(* IEC 61131-3 sources: Digital-Twin/picode/digital-twin-device/openPLC_v3/webserver/st_files (part 2) *)

(* ---- 924959.st ---- *)
TYPE
  datatype0 : BOOL;
END_TYPE

PROGRAM my_first_program
  VAR
    temp AT %IW1.0 : INT;
    out AT %QW0.0 : INT;
  END_VAR
  VAR
    sp : REAL := 1376.0;
    x0 : REAL := 0.0;
    tr : REAL := 0.001;
    td : REAL := 50.0;
    kp : REAL := 0.00005;
    PID0 : PID;
    GT39_OUT : BOOL;
    INT_TO_REAL28_OUT : REAL;
    REAL_TO_INT34_OUT : INT;
  END_VAR

  GT39_OUT := GT(temp, 1200);
  INT_TO_REAL28_OUT := INT_TO_REAL(temp);
  PID0(AUTO := GT39_OUT, PV := INT_TO_REAL28_OUT, SP := sp, X0 := x0, KP := kp, TR := tr, TD := td, CYCLE := T#1s);
  REAL_TO_INT34_OUT := REAL_TO_INT(PID0.XOUT);
  out := REAL_TO_INT34_OUT;
END_PROGRAM

CONFIGURATION Config0

  RESOURCE Res0 ON PLC
    TASK mytask(INTERVAL := T#50ms,PRIORITY := 0);
    PROGRAM my WITH mytask : my_first_program;
  END_RESOURCE
END_CONFIGURATION

(* ---- 925603.st ---- *)
TYPE
  datatype0 : BOOL;
END_TYPE

PROGRAM my_first_program
  VAR
    temp AT %IW1.0 : INT;
    out AT %QW0.0 : INT;
  END_VAR
  VAR
    sp : REAL := 1030.0;
    x0 : REAL := 0.0;
    tr : REAL := 0.001;
    td : REAL := 50.0;
    kp : REAL := 0.00005;
    PID0 : PID;
    GT39_OUT : BOOL;
    INT_TO_REAL28_OUT : REAL;
    REAL_TO_INT34_OUT : INT;
  END_VAR

  GT39_OUT := GT(temp, 1040);
  INT_TO_REAL28_OUT := INT_TO_REAL(temp);
  PID0(AUTO := GT39_OUT, PV := INT_TO_REAL28_OUT, SP := sp, X0 := x0, KP := kp, TR := tr, TD := td, CYCLE := T#1s);
  REAL_TO_INT34_OUT := REAL_TO_INT(PID0.XOUT);
  out := REAL_TO_INT34_OUT;
END_PROGRAM

CONFIGURATION Config0

  RESOURCE Res0 ON PLC
    TASK mytask(INTERVAL := T#50ms,PRIORITY := 0);
    PROGRAM my WITH mytask : my_first_program;
  END_RESOURCE
END_CONFIGURATION

(* ---- 926092.st ---- *)
PROGRAM my_first_program
  VAR
    temp AT %IW0.0 : INT;
    lamp AT %QX0.0 : BOOL;
    lamp1 AT %QX0.2 : BOOL;
  END_VAR
  VAR
    GT7_OUT : BOOL;
    GT1_OUT : BOOL;
  END_VAR

  GT7_OUT := GT(temp, 17170);
  lamp := GT7_OUT;
  GT1_OUT := GT(temp, 18350);
  lamp1 := GT1_OUT;
END_PROGRAM

CONFIGURATION Config0

  RESOURCE Res0 ON PLC
    TASK mytask(INTERVAL := T#50ms,PRIORITY := 0);
    PROGRAM my WITH mytask : my_first_program;
  END_RESOURCE
END_CONFIGURATION

(* ---- 939656.st ---- *)
PROGRAM my_first_program
  VAR
    temp AT %IW0.0 : INT;
    lamp AT %QX0.0 : BOOL;
    lamp1 AT %QX0.2 : BOOL;
  END_VAR
  VAR
    GT7_OUT : BOOL;
    GT1_OUT : BOOL;
  END_VAR

  GT7_OUT := GT(temp, 17170);
  lamp := GT7_OUT;
  GT1_OUT := GT(temp, 18350);
  lamp1 := GT1_OUT;
END_PROGRAM

CONFIGURATION Config0

  RESOURCE Res0 ON PLC
    TASK mytask(INTERVAL := T#50ms,PRIORITY := 0);
    PROGRAM my WITH mytask : my_first_program;
  END_RESOURCE
END_CONFIGURATION

(* ---- 953895.st ---- *)
PROGRAM program0
  VAR
    PID0 : PID;
    Kp : REAL := 0.01;
    Ki : REAL := 0.1;
    Kd : REAL := 50.0;
  END_VAR
  VAR
    Temperature AT %IW1 : UINT;
    Flow AT %QW0 : UINT;
  END_VAR
  VAR
    Setpoint : UINT := 2500;
    Zero : REAL := 0.0;
    GT13_OUT : BOOL;
    UINT_TO_REAL1_OUT : REAL;
    UINT_TO_REAL9_OUT : REAL;
    REAL_TO_UINT11_OUT : UINT;
  END_VAR

  GT13_OUT := GT(Temperature, Setpoint);
  UINT_TO_REAL1_OUT := UINT_TO_REAL(Temperature);
  UINT_TO_REAL9_OUT := UINT_TO_REAL(Setpoint);
  PID0(AUTO := GT13_OUT, PV := UINT_TO_REAL1_OUT, SP := UINT_TO_REAL9_OUT, X0 := Zero, KP := Kp, TR := Ki, TD := Kd, CYCLE := T#50ms);
  REAL_TO_UINT11_OUT := REAL_TO_UINT(PID0.XOUT);
  Flow := REAL_TO_UINT11_OUT;
END_PROGRAM

CONFIGURATION Config0

  RESOURCE Res0 ON PLC
    TASK task0(INTERVAL := T#50ms,PRIORITY := 0);
    PROGRAM instance0 WITH task0 : program0;
  END_RESOURCE
END_CONFIGURATION

(* ---- 966953.st ---- *)
PROGRAM program0
  VAR
    PID0 : PID;
    Kp : REAL := 0.0001;
    Ki : REAL := 0.1;
    Kd : REAL := 50.0;
  END_VAR
  VAR
    Temperature AT %IW0 : UINT;
    Flow AT %QW0 : UINT;
  END_VAR
  VAR
    Setpoint : UINT := 26214;
    Zero : REAL := 0.0;
    GT13_OUT : BOOL;
    UINT_TO_REAL1_OUT : REAL;
    UINT_TO_REAL9_OUT : REAL;
    REAL_TO_UINT11_OUT : UINT;
  END_VAR

  GT13_OUT := GT(Temperature, Setpoint);
  UINT_TO_REAL1_OUT := UINT_TO_REAL(Temperature);
  UINT_TO_REAL9_OUT := UINT_TO_REAL(Setpoint);
  PID0(AUTO := GT13_OUT, PV := UINT_TO_REAL1_OUT, SP := UINT_TO_REAL9_OUT, X0 := Zero, KP := Kp, TR := Ki, TD := Kd, CYCLE := T#50ms);
  REAL_TO_UINT11_OUT := REAL_TO_UINT(PID0.XOUT);
  Flow := REAL_TO_UINT11_OUT;
END_PROGRAM

CONFIGURATION Config0

  RESOURCE Res0 ON PLC
    TASK task0(INTERVAL := T#50ms,PRIORITY := 0);
    PROGRAM instance0 WITH task0 : program0;
  END_RESOURCE
END_CONFIGURATION

(* ---- 970422.st ---- *)
PROGRAM my_first_program
  VAR
    temp AT %IW0.0 : INT;
    out AT %QW0.0 : INT;
  END_VAR
  VAR
    sp : REAL := 2293.0;
    x0 : REAL := 0.0;
    tr : REAL := 1.0;
    td : REAL := 1.0;
    kp : REAL := 2.0;
    PID0 : PID;
    INT_TO_REAL28_OUT : REAL;
    REAL_TO_INT32_OUT : INT;
  END_VAR

  INT_TO_REAL28_OUT := INT_TO_REAL(temp);
  PID0(AUTO := TRUE, PV := INT_TO_REAL28_OUT, SP := sp, X0 := x0, KP := kp, TR := tr, TD := td, CYCLE := T#1s);
  REAL_TO_INT32_OUT := REAL_TO_INT(PID0.XOUT);
  out := REAL_TO_INT32_OUT;
END_PROGRAM

CONFIGURATION Config0

  RESOURCE Res0 ON PLC
    TASK mytask(INTERVAL := T#50ms,PRIORITY := 0);
    PROGRAM my WITH mytask : my_first_program;
  END_RESOURCE
END_CONFIGURATION

(* ---- 979458.st ---- *)
PROGRAM my_first_program
  VAR
    temp AT %IW0.0 : INT;
    out AT %QW0.0 : INT;
  END_VAR
  VAR
    sp : REAL := 2500.0;
    x0 : REAL := 0.0;
    tr : REAL := 0.1;
    td : REAL := 50.0;
    kp : REAL := 0.01;
    PID0 : PID;
    INT_TO_REAL28_OUT : REAL;
    REAL_TO_INT34_OUT : INT;
  END_VAR

  INT_TO_REAL28_OUT := INT_TO_REAL(temp);
  PID0(AUTO := TRUE, PV := INT_TO_REAL28_OUT, SP := sp, X0 := x0, KP := kp, TR := tr, TD := td, CYCLE := T#1s);
  REAL_TO_INT34_OUT := REAL_TO_INT(PID0.XOUT);
  out := REAL_TO_INT34_OUT;
END_PROGRAM

CONFIGURATION Config0

  RESOURCE Res0 ON PLC
    TASK mytask(INTERVAL := T#50ms,PRIORITY := 0);
    PROGRAM my WITH mytask : my_first_program;
  END_RESOURCE
END_CONFIGURATION

(* ---- 980664.st ---- *)
PROGRAM my_first_program
  VAR
    temp AT %IW0.0 : INT;
    out AT %QW0.0 : INT;
  END_VAR
  VAR
    sp : REAL := 1930.0;
    x0 : REAL := 0.0;
    tr : REAL := 0.001;
    td : REAL := 50.0;
    kp : REAL := 0.0007;
    PID0 : PID;
    GT36_OUT : BOOL;
    INT_TO_REAL28_OUT : REAL;
    REAL_TO_INT34_OUT : INT;
  END_VAR

  GT36_OUT := GT(temp, 1700);
  INT_TO_REAL28_OUT := INT_TO_REAL(temp);
  PID0(AUTO := GT36_OUT, PV := INT_TO_REAL28_OUT, SP := sp, X0 := x0, KP := kp, TR := tr, TD := td, CYCLE := T#1s);
  REAL_TO_INT34_OUT := REAL_TO_INT(PID0.XOUT);
  out := REAL_TO_INT34_OUT;
END_PROGRAM

CONFIGURATION Config0

  RESOURCE Res0 ON PLC
    TASK mytask(INTERVAL := T#50ms,PRIORITY := 0);
    PROGRAM my WITH mytask : my_first_program;
  END_RESOURCE
END_CONFIGURATION

(* ---- 982831.st ---- *)
TYPE
  datatype0 : BOOL;
END_TYPE

PROGRAM my_first_program
  VAR
    temp AT %IW0.0 : INT;
    out AT %QW0.0 : INT;
  END_VAR
  VAR
    sp : REAL := 2140.0;
    x0 : REAL := 0.0;
    tr : REAL := 0.0006;
    td : REAL := 50.0;
    kp : REAL := 0.0001;
    PID0 : PID;
    INT_TO_REAL28_OUT : REAL;
    REAL_TO_INT34_OUT : INT;
  END_VAR

  INT_TO_REAL28_OUT := INT_TO_REAL(temp);
  PID0(AUTO := TRUE, PV := INT_TO_REAL28_OUT, SP := sp, X0 := x0, KP := kp, TR := tr, TD := td, CYCLE := T#1s);
  REAL_TO_INT34_OUT := REAL_TO_INT(PID0.XOUT);
  out := REAL_TO_INT34_OUT;
END_PROGRAM

CONFIGURATION Config0

  RESOURCE Res0 ON PLC
    TASK mytask(INTERVAL := T#50ms,PRIORITY := 0);
    PROGRAM my WITH mytask : my_first_program;
  END_RESOURCE
END_CONFIGURATION

(* ---- 983137.st ---- *)
TYPE
  datatype0 : BOOL;
END_TYPE

PROGRAM my_first_program
  VAR
    temp AT %IW1.0 : INT;
    out AT %QW0.0 : INT;
  END_VAR
  VAR
    sp : REAL := 1030.0;
    x0 : REAL := 0.0;
    tr : REAL := 0.001;
    td : REAL := 50.0;
    kp : REAL := 0.00005;
    PID0 : PID;
    GT39_OUT : BOOL;
    INT_TO_REAL28_OUT : REAL;
    REAL_TO_INT34_OUT : INT;
  END_VAR

  GT39_OUT := GT(temp, 950);
  INT_TO_REAL28_OUT := INT_TO_REAL(temp);
  PID0(AUTO := GT39_OUT, PV := INT_TO_REAL28_OUT, SP := sp, X0 := x0, KP := kp, TR := tr, TD := td, CYCLE := T#1s);
  REAL_TO_INT34_OUT := REAL_TO_INT(PID0.XOUT);
  out := REAL_TO_INT34_OUT;
END_PROGRAM

CONFIGURATION Config0

  RESOURCE Res0 ON PLC
    TASK mytask(INTERVAL := T#50ms,PRIORITY := 0);
    PROGRAM my WITH mytask : my_first_program;
  END_RESOURCE
END_CONFIGURATION

(* ---- blank_program.st ---- *)
PROGRAM prog0
  VAR
    var_in : BOOL;
    var_out : BOOL;
  END_VAR

  var_out := var_in;
END_PROGRAM

CONFIGURATION Config0

  RESOURCE Res0 ON PLC
    TASK Main(INTERVAL := T#50ms,PRIORITY := 0);
    PROGRAM Inst0 WITH Main : prog0;
  END_RESOURCE
END_CONFIGURATION
